(* KBO coating-state enum. UINT-typed so REFERENCE TO E_KBO_CoatingStates
   is bridge-compatible with the ND mover's REFERENCE TO UINT. *)
{attribute 'qualified_only'}
{attribute 'strict'}
TYPE E_KBO_CoatingStates :
(
    Unknown := 0,
    Si := 1,
    B4C := 2
) UINT;
END_TYPE

(* stored: Version 1.1.0.1
   DUT E_KBO_CoatingStates: Id {a3f1b2c4-5d6e-47f8-9a0b-1c2d3e4f5a6b} *)
